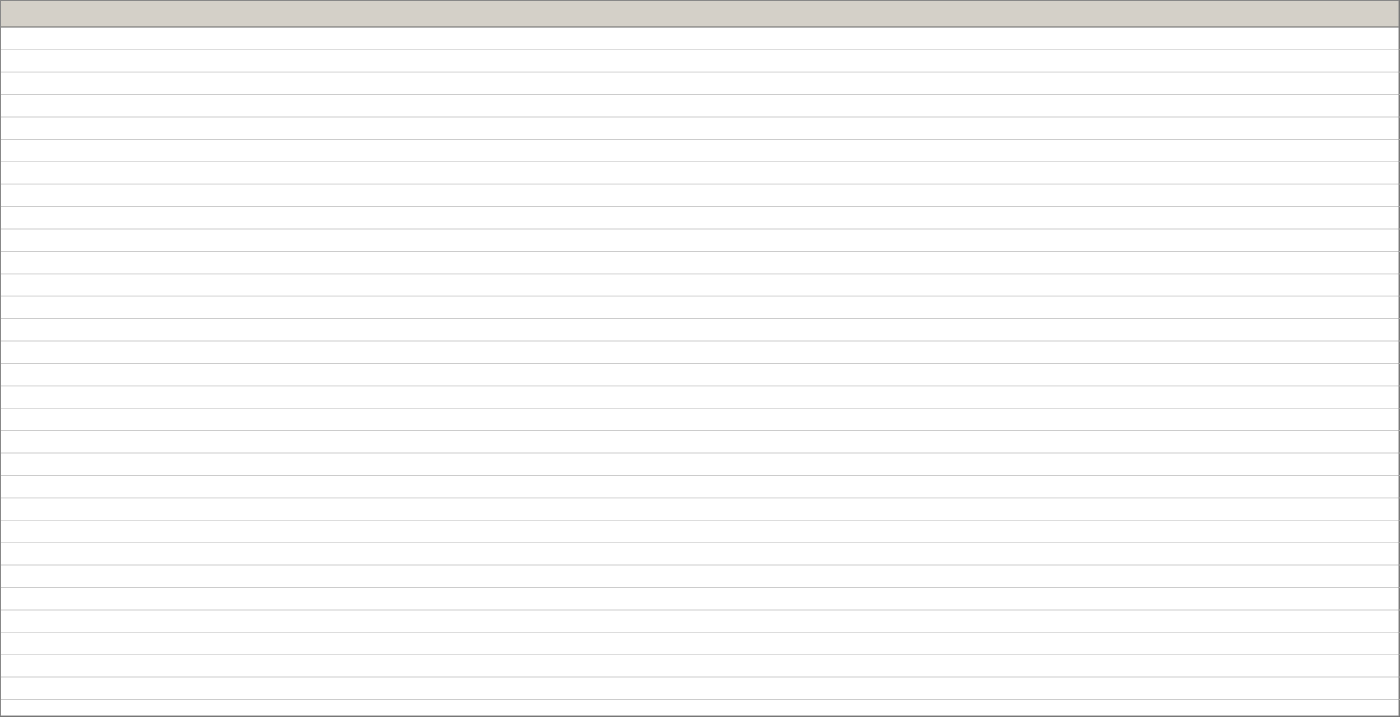
VISUALIZATION vis_Error_History  // 1560x800
    Table (0,0 1560x800), data array: Buffer_Act_History
        p3854506369: Buffer_Act_History[INDEX].sDateTime
        p1892666644: Buffer_Act_History[INDEX].sErrID
        p338671338: Buffer_Act_History[INDEX].sLevel
        p2170511999: Buffer_Act_History[INDEX].sModuleDescription
        p3723444502: Buffer_Act_History[INDEX].sErrorMessage
        p4092479075: Module Description
        p2237128397: Error Message
END_VISUALIZATION

(* stored: Version 1.1.0.1, ProductVersion 3.1.4024.13
   Visu vis_Error_History: Id {660f19fe-0831-4045-9aeb-8c8cf2775605} *)
